Fanuc KAREL source: kb00076.KL

PROGRAM KB00076
%STACKSIZE=65535
%PRIORITY=65535
%NOLOCKGROUP
VAR
P1 : POSITION
P2 : POSITION
P3 : POSITION
RESULT : POSITION
BEGIN
-- UNRESOLVED_PC line 9 opcodes [27 22 1C 22 1C 22 1C 76 7E 4A] marker_code=0
END KB00076
